(* IEC 61131-3 sources: plc-process-lib/src/POUs/PRG_Main, 1 file *)

(* ---- PRG_Main.decl.st ---- *)
// Назначение: служебная программа рабочей сборки (cds.py build, режим normal), не часть API
//             библиотеки. CODESYS 3.5.17 не собирает приложение с пустой конфигурацией задач
//             («Не задано ни одной задачи»), а cds.py всегда создаёт её, поэтому задаче MainTask
//             нужна программа. Единственное действие — показать системное время библиотеки для
//             ручной проверки монотонности LTIME() онлайн (R1, docs/MANUAL_STEPS.md). Компилятор
//             проверяет только объекты, достижимые из задач, поэтому проверку всех объектов
//             библиотеки даёт тестовая сборка (cds.py build --tests, cds.py test).
//             В .library программа не входит.
// Автор:      kr0nsch
// Версия:     0.1.0
// Документ:   docs/ASSUMPTIONS.md, решения F-02 и F-03
PROGRAM PRG_Main
VAR
    fbSysTime : FB_SystemTime;   // системный источник времени библиотеки
    ltUptime  : LTIME;           // время от старта рантайма (оператор LTIME()), для онлайн-просмотра
END_VAR
